Universal Robots URScript: T009_mistralai_Mistral-Large-3-675B-Instruct-2512-NVFP4_edit_perf_rep1.urscript

# Task: T009 — Laser surface scan — fenced mode (Optimized)
# Optimized for faster cycle time while maintaining safety constraints

def task_T009():
  TCP_SPEED_CAP = 0.200
  def safe_movel(pose, a, v, r):
    movel(pose, a=a, v=min(v, TCP_SPEED_CAP), r=r)
  end

  # [0] Verify E-Stop
  if (get_digital_in(0) == True):
    popup("E-Stop active — aborting program.", error=True)
    halt
  end

  # [1] Home - Increased speed and acceleration
  movej([0.0000, -1.5708, 1.5708, -1.5708, -1.5708, 0.0000], a=2.0000, v=1.0000)

  # [2] Above scan start - Increased speed
  safe_movel(p[0.250000, -0.100000, 0.250000, 0.0000, 3.1416, 0.0000], 1.2000, 0.2000, 0.0100)

  # [3] Descend to scan height - Increased speed
  safe_movel(p[0.250000, -0.100000, 0.120000, 0.0000, 3.1416, 0.0000], 0.8000, 0.1500, 0.0050)

  # [4] Laser ON
  set_digital_out(3, True)

  # [5] Scan line 1 - Increased acceleration
  safe_movel(p[0.250000, 0.100000, 0.120000, 0.0000, 3.1416, 0.0000], 0.5000, 0.0500, 0.0050)

  # [6] Step to line 2 - Increased speed and acceleration
  safe_movel(p[0.350000, 0.100000, 0.120000, 0.0000, 3.1416, 0.0000], 0.8000, 0.1500, 0.0050)

  # [7] Scan line 2 reverse - Increased acceleration
  safe_movel(p[0.350000, -0.100000, 0.120000, 0.0000, 3.1416, 0.0000], 0.5000, 0.0500, 0.0050)

  # [8] Step to line 3 - Increased speed and acceleration
  safe_movel(p[0.450000, -0.100000, 0.120000, 0.0000, 3.1416, 0.0000], 0.8000, 0.1500, 0.0050)

  # [9] Scan line 3 - Increased acceleration
  safe_movel(p[0.450000, 0.100000, 0.120000, 0.0000, 3.1416, 0.0000], 0.5000, 0.0500, 0.0050)

  # [10] Step to line 4 - Increased speed and acceleration
  safe_movel(p[0.550000, 0.100000, 0.120000, 0.0000, 3.1416, 0.0000], 0.8000, 0.1500, 0.0050)

  # [11] Scan line 4 reverse - Increased acceleration, removed blend radius
  safe_movel(p[0.550000, -0.100000, 0.120000, 0.0000, 3.1416, 0.0000], 0.5000, 0.0500, 0.0)

  # [12] Laser OFF
  set_digital_out(3, False)

  # [13] Retract - Increased speed
  safe_movel(p[0.400000, 0.000000, 0.300000, 0.0000, 3.1416, 0.0000], 1.2000, 0.2000, 0.0100)

  # [14] Return home - Increased speed and acceleration
  movej([0.0000, -1.5708, 1.5708, -1.5708, -1.5708, 0.0000], a=2.0000, v=1.0000)
end

# Entry point
task_T009()
